// Type d'une variable (docs/06 § 2)
{attribute 'qualified_only'}
{attribute 'strict'}
TYPE E_VarType :
(
    Number := 0,
    Bool := 1,
    Position := 2
) USINT;
END_TYPE

(* stored: Version 1.1.0.1, ProductVersion 3.1.4024.12
   DUT E_VarType: Id {ea41ac98-963f-5f84-b064-7d6112c80e04} *)
